Staubli VAL3: loadLib.pgx

public program loadLib(num x_nLib, num& x_nResult)
  local string l_sPath
begin
  if x_nLib>=0
    l_sPath="Disk://data/CustomerLib/lib"+toString("",x_nLib)+"/safeData"
    x_nResult=safeData:libLoad(l_sPath)
    wait(x_nResult==0)
  else
    call rs:setAlarm(302,0)
  endIf
end
